TYPE ST_PolarIIChamber_ArmRotateServiceStatus :
STRUCT
	JogPositive : ST_ServiceStatus;
	JogNegative : ST_ServiceStatus;
	IncrementalJog : ST_ServiceStatus;
	MoveRecipe : ST_ServiceStatus;
	NegLimitPos : ST_ServiceStatus;
	PosLimitPos : ST_ServiceStatus;
	NozzlePortPos : ST_ServiceStatus;
	Noz1CenterPos : ST_ServiceStatus;
	Noz2CenterPos : ST_ServiceStatus;
	Noz3CenterPos : ST_ServiceStatus;
END_STRUCT
END_TYPE

(* stored: Version 1.1.0.1, ProductVersion 3.1.4026.18
   DUT ST_PolarIIChamber_ArmRotateServiceStatus: Id {14000000-0000-0000-0000-000000000027} *)
